FUNCTION FC 1 : VOID
BEGIN
NETWORK
END_ORGANIZATION_BLOCK
